// TIA Portal V17 export
ORGANIZATION_BLOCK "Main"   // OB1, LAD, ProgramCycle
TITLE = Programa principal
{ S7_Optimized_Access := 'TRUE' }
// Generado automáticamente con Claude Code + TIA Openness
   VAR_INPUT
      Initial_Call : Bool;   // Initial call of this OB
      Remanence : Bool;   // =True, if remanent data are available
   END_VAR
BEGIN

REGION Network 1: Motor 1
   // Llamada al bloque de arranque y paro con las entradas/salidas físicas
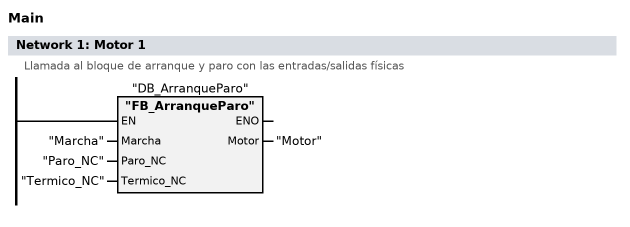
   RUNG wire#powerrail
      "DB_ArranqueParo"(Marcha := "Marcha", Paro_NC := "Paro_NC", Termico_NC := "Termico_NC", Motor => "Motor")
   END_RUNG
   // the same network as SCL:
   "DB_ArranqueParo"(Marcha := "Marcha", Paro_NC := "Paro_NC", Termico_NC := "Termico_NC", Motor => "Motor");   // "FB_ArranqueParo"
END_REGION
END_ORGANIZATION_BLOCK
